(* CODESYS project PROV9.project

Project tree, tasks and I/O mapping:
  Device : CODESYS Control Win V3, 3S - Smart Software Solutions GmbH, order no. 305021, version 3.5.9.10
    application Application
      libraries: Standard, * (System)
      task MainTask (cyclic, interval t#20ms, priority 1) calls PLC_PRG, VARIABLES, M_TIEMPOS, SENSOR_P, SENSOR_C
      program PLC_PRG [LD]
      global variables GVL
      Symbols
      program VARIABLES [ST]
      program EM [ST]
      program M_TIEMPOS [ST]
      program EA [ST]
      program SENSOR_P [ST]
      data type U_REAL_WORDS
      program SENSOR_C [ST]
    Ethernet : Ethernet, 3S - Smart Software Solutions GmbH, version 3.5.15.0
        settings: IPAddress = [10,20,64,7]; SubnetMask = [255,255,255,0]; GatewayAddress = [10,20,64,1]; MACAddress = [16#DC,16#46,16#28,16#0A,16#44,16#B1]; NetworkInterfaceName = 'Wi-Fi'; NetworkInterfaceName = "Wi-Fi"; SaveCommunicationSettings = FALSE
      Modbus_TCP_Master : Modbus TCP Master, 3S - Smart Software Solutions GmbH, version 3.5.15.0
        Modbus_TCP_Slave : Modbus TCP Slave, 3S - Smart Software Solutions GmbH, version 3.5.15.0
            settings: Unit-ID = 1; IPAddress = [192, 168, 10, 24]; Port = 5020; COMANDO.Function Code = 6; COMANDO.Read Offset = 0; COMANDO.Read Length = 0; COMANDO.Write Offset = 16#0000; COMANDO.Write Length = 1; COMANDO.Cycle Time = 100; CONFIRMACION.Function Code = 3; CONFIRMACION.Read Offset = 16#0001; CONFIRMACION.Read Length = 1; CONFIRMACION.Write Offset = 0; CONFIRMACION.Write Length = 0; CONFIRMACION.Cycle Time = 100
            output Application.CONFIRMACION : WORD  // COMANDO
            input  Application.COMANDO : WORD  // CONFIRMACION
      ModbusTCP_Slave_Device : ModbusTCP Slave Device, 3S - Smart Software Solutions GmbH, version 3.5.15.0
          input  Application.CONFIRMACION : WORD  // Inputs.Inputs
          output Application.COMANDO : WORD  // Outputs.Outputs
          output Application.TIEMPO_AP_MOD : WORD  // Outputs.Outputs
          output Application.TIEMPO_AN_MOD : WORD  // Outputs.Outputs
          output Application.TIEMPO_BP_MOD : WORD  // Outputs.Outputs
          output Application.TIEMPO_BN_MOD : WORD  // Outputs.Outputs
          output Application.TIEMPO_CP_MOD : WORD  // Outputs.Outputs
          output Application.TIEMPO_CN_MOD : WORD  // Outputs.Outputs
          output Application.CICLO_ACTUAL : WORD  // Outputs.Outputs
          output Application.PresionWord0 : WORD  // Outputs.Outputs
          output Application.PresionWord1 : WORD  // Outputs.Outputs
          output Application.CaudalPromedioWord0 : WORD  // Outputs.Outputs
          output Application.CaudalPromedioWord1 : WORD  // Outputs.Outputs
          unmapped channels: Inputs, Outputs
*)

// Device/Application/U_REAL_WORDS
TYPE U_REAL_WORDS :
UNION
    RealValue : REAL;
    Words : ARRAY[0..1] OF WORD;
END_UNION
END_TYPE

// Device/Application/GVL
VAR_GLOBAL
	IN0:BYTE;
	OUT0:BYTE;
	IN1:BYTE;
	OUT1:BYTE;
	FIN_CICLO:BOOL;
	
	// VARIABLES //
	START:BOOL;
	START_A: BOOL;
	STOP:BOOL;
	AN:BOOL;
	AP:BOOL;
	BN:BOOL;
	BP:BOOL;
	CN:BOOL;
	CP:BOOL;
	SP:BOOL; // SENSOR CAJAS
	
	// SENSORES ANALOGOS
	PRESION_V: REAL;
	PRESION: REAL;
	PresionModbus : U_REAL_WORDS;
    PresionWord0 : WORD;
    PresionWord1 : WORD;
	
	
    // AUTOTESTING: CAUDAL PROMEDIO
	CAUDAL_V: REAL;
	CAUDAL: REAL;
    SUMA_CAUDAL : LREAL := 0.0;
    CONTADOR_CAUDAL : UDINT := 0;
    CAUDAL_PROMEDIO_CICLO : REAL := 0.0;
    CAUDAL_PROMEDIO_LISTO : BOOL := FALSE;
    MEDIR_CAUDAL : BOOL := FALSE;
    CICLO_FIN_PROCESADO : BOOL := FALSE;
	
    // PROMEDIO DE CAUDAL PARA MODBUS
    CaudalPromedioModbus : U_REAL_WORDS;
    CaudalPromedioWord0 : WORD;
    CaudalPromedioWord1 : WORD;



	


	CONFIRMACION:WORD;
	COMANDO:WORD:=456;
	
	//OUT
	MAP:BOOL;
	MAN:BOOL;
	MBP:BOOL;
	MBN:BOOL;
	MCP:BOOL; //ECECTROVALVULA MONO ESTABLE
	LEDV:BOOL;
	LEDA:BOOL;
	LEDR:BOOL;
	BUZZER:BOOL; //SIRENA
	
	// TIEMPOS DE CILINDROS

	TIEMPO_AP_MOD : WORD;
	TIEMPO_AN_MOD : WORD;

	TIEMPO_BP_MOD : WORD;
	TIEMPO_BN_MOD : WORD;

	TIEMPO_CP_MOD : WORD;
	TIEMPO_CN_MOD : WORD;

	CICLO_ACTUAL : UINT;
	FIN_CICLO_MB:WORD;
	
END_VAR

// Device/Application/PLC_PRG
PROGRAM PLC_PRG
VAR
	M0: BOOL;
	M1: BOOL;
END_VAR
VAR // added by the converter: edge detectors and wires of the graphical bodies
    _w1, _w2 : BOOL;
END_VAR

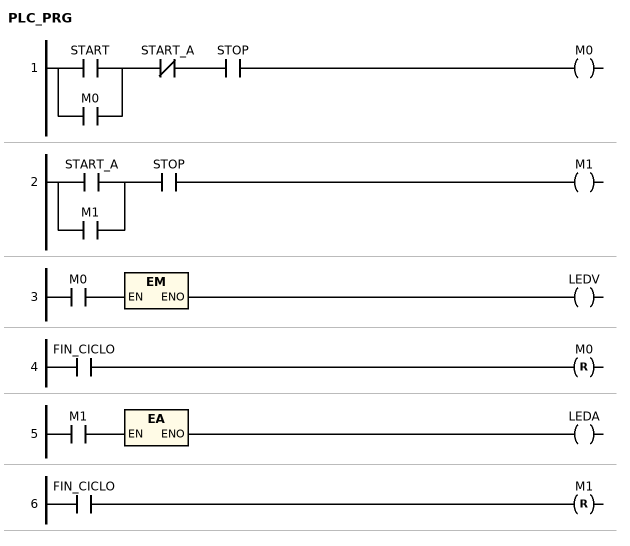
// NETWORK 1
M0 := (START OR M0) AND NOT START_A AND STOP;

// NETWORK 2
M1 := (START_A OR M1) AND STOP;

// NETWORK 3
_w1 := M0;
IF _w1 THEN EM(); END_IF
LEDV := _w1;

// NETWORK 4
M0 R= FIN_CICLO;

// NETWORK 5
_w2 := M1;
IF _w2 THEN EA(); END_IF
LEDA := _w2;

// NETWORK 6
M1 R= FIN_CICLO;

END_PROGRAM

// Device/Application/EM
PROGRAM EM
VAR
	T0:TON;
	T10:TON;
	T20:TON;
	T30:TON;
	T40:TON;
	T50:TON;
	T60:TON;
	T70:TON;
	T80:TON;
	T90:TON;
	
	VP:INT;
END_VAR

CASE VP OF
	0:
		FIN_CICLO:=FALSE;
		T50(IN:=FALSE);
		T0(IN:=TRUE, PT:=T#200MS);
		IF PLC_PRG.M0 AND SP AND AN AND BN AND CN AND T0.Q THEN
			MAP:=TRUE;
			VP:=10;
		END_IF
	
	10:
		T0(IN:=FALSE);
		T10(IN:=TRUE, PT:=T#200MS);
		IF AP AND BN AND CN AND T10.Q THEN
			MBP:=TRUE;
			VP:=20;
		END_IF
		
	20:
		T10(IN:=FALSE);
		T20(IN:=TRUE, PT:=T#500MS);
		IF AP AND BP AND CN AND T20.Q THEN
			MBP:=FALSE;
			MBN:=TRUE;
			VP:=30;
		END_IF
		
	30:
		T20(IN:=FALSE);
		T30(IN:=TRUE, PT:=T#200MS);
		IF AP AND BN AND CN AND T30.Q THEN
			MAP:=FALSE;
			MAN:=TRUE;
			VP:=40;
		END_IF
		
	40:
		T30(IN:=FALSE);
		T40(IN:=TRUE, PT:=T#200MS);
		IF AN AND BN AND CN AND T40.Q THEN
			MCP:=TRUE;
			VP:=50;
		END_IF
		
	50:
		T40(IN:=FALSE);
		T50(IN:=TRUE, PT:=T#200MS);
		IF AN AND BN AND CP AND T50.Q THEN
			FIN_CICLO:=TRUE;
			MCP:=FALSE;
			MAN:=FALSE;
			MBN:=FALSE;
			VP:=0;
		END_IF
		
END_CASE

END_PROGRAM

// Device/Application/EA
PROGRAM EA
VAR
	T0:TON;
	T10:TON;
	T20:TON;
	T30:TON;
	T40:TON;
	T50:TON;
	T60:TON;
	T70:TON;
	T80:TON;
	T90:TON;
	T_FIN : TON;
	VP:INT;
END_VAR

CASE VP OF
	0:
		T_FIN(IN:=FALSE);
		FIN_CICLO:=FALSE;
		T50(IN:=FALSE);
		T0(IN:=TRUE, PT:=T#200MS);
		IF PLC_PRG.M1 AND AN AND BN AND CN AND T0.Q THEN
			MAP:=TRUE;
			VP:=10;
		END_IF
	
	10:
		T0(IN:=FALSE);
		T10(IN:=TRUE, PT:=T#200MS);
		IF AP AND BN AND CN AND T10.Q THEN
			MBP:=TRUE;
			VP:=20;
		END_IF
		
	20:
		T10(IN:=FALSE);
		T20(IN:=TRUE, PT:=T#500MS);
		IF AP AND BP AND CN AND T20.Q THEN
			MBP:=FALSE;
			MBN:=TRUE;
			VP:=30;
		END_IF
		
	30:
		T20(IN:=FALSE);
		T30(IN:=TRUE, PT:=T#200MS);
		IF AP AND BN AND CN AND T30.Q THEN
			MAP:=FALSE;
			MAN:=TRUE;
			VP:=40;
		END_IF
		
	40:
		T30(IN:=FALSE);
		T40(IN:=TRUE, PT:=T#200MS);
		IF AN AND BN AND CN AND T40.Q THEN
			MCP:=TRUE;
			VP:=50;
		END_IF
		
	50:
		T40(IN:=FALSE);
		T50(IN:=TRUE, PT:=T#200MS);
		IF AN AND BN AND CP AND T50.Q THEN
			FIN_CICLO:=TRUE;
			MCP:=FALSE;
			MAN:=FALSE;
			MBN:=FALSE;
			
			VP:=60;
		END_IF
		
	60:
    T50(IN:=FALSE);
    T_FIN(IN:=TRUE, PT:=T#3S);

    IF T_FIN.Q THEN
        VP := 0;
    END_IF
		
END_CASE

END_PROGRAM

// Device/Application/VARIABLES
PROGRAM VARIABLES
VAR
END_VAR

START:=IN0.0;
STOP:=IN0.1;
START_A:=IN1.1;
AN:=IN0.2;
AP:=IN0.3;
BN:=IN0.4;
BP:=IN0.5;
CN:=IN0.6;
CP:=IN0.7;
SP:=IN1.0;

OUT0.0:=MAP;
OUT0.1:=MAN;
OUT0.2:=MBP;
OUT0.3:=MBN;
OUT0.4:=MCP;
OUT0.5:=LEDV;
OUT0.6:=LEDA;
OUT0.7:=LEDR;
OUT1.0:=BUZZER;

END_PROGRAM

// Device/Application/M_TIEMPOS
PROGRAM M_TIEMPOS
VAR
    // Temporizadores de medición
    T_AP : TON;
	T_AN : TON;
    T_BP : TON;
    T_BN : TON;
    T_CP : TON;
    T_CN : TON;

    // Tiempos medidos
    Tiempo_AP : TIME;
	Tiempo_AN : TIME;
    Tiempo_BP : TIME;
    Tiempo_BN : TIME;
    Tiempo_CP : TIME;
    Tiempo_CN : TIME;

    // Banderas para indicar que se está midiendo
    Ciclo_Completo : BOOL;
	Numero_Ciclo : UINT;
	Medir_AP : BOOL;
	Medir_AN : BOOL;
    Medir_BP : BOOL;
    Medir_BN : BOOL;
    Medir_CP : BOOL;
    Medir_CN : BOOL;
END_VAR

// =====================================================
// TEMPORIZADORES
// =====================================================

T_AP(
    IN := Medir_AP,
    PT := T#10S
);

T_BP(
    IN := Medir_BP,
    PT := T#10S
);

T_BN(
    IN := Medir_BN,
    PT := T#10S
);

T_AN(
    IN := Medir_AN,
    PT := T#10S
);

T_CP(
    IN := Medir_CP,
    PT := T#10S
);

T_CN(
    IN := Medir_CN,
    PT := T#10S
);


// =====================================================
// CICLO COMPLETO
// =====================================================

Ciclo_Completo := FALSE;


// =====================================================
// A+
// MAP → AP
// =====================================================

IF MAP AND NOT AP AND NOT Medir_AP THEN
    Medir_AP := TRUE;
END_IF;

IF AP AND Medir_AP THEN
    Tiempo_AP := T_AP.ET;
    Medir_AP := FALSE;
END_IF;


// =====================================================
// B+
// MBP → BP
// =====================================================

IF MBP AND NOT BP AND NOT Medir_BP THEN
    Medir_BP := TRUE;
END_IF;

IF BP AND Medir_BP THEN
    Tiempo_BP := T_BP.ET;
    Medir_BP := FALSE;
END_IF;


// =====================================================
// B-
// MBN → BN
// =====================================================

IF MBN AND NOT BN AND NOT Medir_BN THEN
    Medir_BN := TRUE;
END_IF;

IF BN AND Medir_BN THEN
    Tiempo_BN := T_BN.ET;
    Medir_BN := FALSE;
END_IF;


// =====================================================
// A-
// MAN → AN
// =====================================================

IF MAN AND NOT AN AND NOT Medir_AN THEN
    Medir_AN := TRUE;
END_IF;

IF AN AND Medir_AN THEN
    Tiempo_AN := T_AN.ET;
    Medir_AN := FALSE;
END_IF;


// =====================================================
// C+
// MCP → CP
// =====================================================

IF MCP AND NOT CP AND NOT Medir_CP THEN
    Medir_CP := TRUE;
END_IF;

IF CP AND Medir_CP THEN
    Tiempo_CP := T_CP.ET;
    Medir_CP := FALSE;
END_IF;


// =====================================================
// C-
// MCP = FALSE → CN
// =====================================================

IF NOT MCP AND CP AND NOT CN AND NOT Medir_CN THEN
    Medir_CN := TRUE;
END_IF;

IF CN AND Medir_CN THEN
    Tiempo_CN := T_CN.ET;
    Medir_CN := FALSE;

    // Se completaron los seis movimientos
	Numero_Ciclo := Numero_Ciclo + 1;
    Ciclo_Completo := TRUE;
END_IF;
// =====================================================
// ENVIO DE TIEMPOS A MODBUS
// =====================================================

TIEMPO_AP_MOD := TIME_TO_WORD(Tiempo_AP);
TIEMPO_AN_MOD := TIME_TO_WORD(Tiempo_AN);

TIEMPO_BP_MOD := TIME_TO_WORD(Tiempo_BP);
TIEMPO_BN_MOD := TIME_TO_WORD(Tiempo_BN);

TIEMPO_CP_MOD := TIME_TO_WORD(Tiempo_CP);
TIEMPO_CN_MOD := TIME_TO_WORD(Tiempo_CN);

CICLO_ACTUAL := Numero_Ciclo;

//FIN DE CICLO
FIN_CICLO := Ciclo_Completo;

IF FIN_CICLO THEN
    FIN_CICLO_MB := 1;
ELSE
    FIN_CICLO_MB := 0;
END_IF;

END_PROGRAM

// Device/Application/SENSOR_P
PROGRAM SENSOR_P
VAR
END_VAR

// PRESIÓN
// 0...32768 RAW = 0...10 V
// 0...10 V = 0...10 bar

PRESION := (PRESION_V * 10.0) / 32768.0;

PresionModbus.RealValue := PRESION;

PresionWord0 := PresionModbus.Words[0];
PresionWord1 := PresionModbus.Words[1];

END_PROGRAM

// Device/Application/SENSOR_C
PROGRAM SENSOR_C

VAR
    TIMER_MUESTREO_CAUDAL : TON;
    TOMAR_MUESTRA_CAUDAL : BOOL := FALSE;
END_VAR


(* CONVERSION DEL CAUDAL INSTANTANEO *)
CAUDAL := (CAUDAL_V * 100.0) / 32768.0;

(* TEMPORIZADOR DE MUESTREO: 100 ms *)
TIMER_MUESTREO_CAUDAL(
    IN := MEDIR_CAUDAL AND NOT TOMAR_MUESTRA_CAUDAL,
    PT := T#100MS
);

TOMAR_MUESTRA_CAUDAL := TIMER_MUESTREO_CAUDAL.Q;

(* INICIAR MEDICION AL COMENZAR EL CICLO *)
IF MAP AND NOT MEDIR_CAUDAL AND NOT FIN_CICLO THEN
    SUMA_CAUDAL := 0.0;
    CONTADOR_CAUDAL := 0;
    CAUDAL_PROMEDIO_LISTO := FALSE;
    CICLO_FIN_PROCESADO := FALSE;
    MEDIR_CAUDAL := TRUE;
END_IF;

(* TOMAR UNA MUESTRA CADA 100 ms *)
IF TOMAR_MUESTRA_CAUDAL
   AND MEDIR_CAUDAL
   AND NOT FIN_CICLO THEN

    SUMA_CAUDAL := SUMA_CAUDAL + REAL_TO_LREAL(CAUDAL);
    CONTADOR_CAUDAL := CONTADOR_CAUDAL + 1;

END_IF;

(* CALCULAR EL PROMEDIO AL FINAL DEL CICLO *)
IF MEDIR_CAUDAL AND FIN_CICLO
   AND NOT CICLO_FIN_PROCESADO THEN

    IF CONTADOR_CAUDAL > 0 THEN
        CAUDAL_PROMEDIO_CICLO :=
            LREAL_TO_REAL(
                SUMA_CAUDAL / UDINT_TO_LREAL(CONTADOR_CAUDAL)
            );

        CAUDAL_PROMEDIO_LISTO := TRUE;
    END_IF;

    MEDIR_CAUDAL := FALSE;
    CICLO_FIN_PROCESADO := TRUE;
END_IF;

(* ENVIAR PROMEDIO DE CAUDAL A MODBUS *)
CaudalPromedioModbus.RealValue := CAUDAL_PROMEDIO_CICLO;

CaudalPromedioWord0 := CaudalPromedioModbus.Words[0];
CaudalPromedioWord1 := CaudalPromedioModbus.Words[1];

END_PROGRAM
